Fanuc KAREL source: KA00169.KL

PROGRAM KA00169
%NOLOCKGROUP
VAR
  SRC: ARRAY[4] OF BOOLEAN
  DST: ARRAY[4] OF VECTOR
BEGIN
  DST = SRC
END KA00169
